Fanuc KAREL source: kd00042.KL

-- PROVISIONAL review KL for V770-1; original PC SHA256 14c779a276e6f473537c1e177adf0885141d48ee65f29f4c4c44e73cbc90e743
-- Incomplete behavior may be omitted. Consult companion uncertainty JSON. Do not deploy.
PROGRAM KD00042
%NOLOCKGROUP
VAR
  I : INTEGER
  J : INTEGER
  B : BOOLEAN
  R : REAL
  S : STRING[80]
-- UNRESOLVED_DECL N type=001100
BEGIN
  -- UNRESOLVED_PC offsets 5-12; opcodes 9D,23
  -- UNRESOLVED_PC offsets 17-21; opcodes 7F
END KD00042
